{attribute 'no_assign'}
FUNCTION_BLOCK FB_DO_WTURBINE_LD0_LPHD1_Proxy EXTENDS FB_AcsiCommonDataClass
VAR_INPUT
	stVal: FB_AcsiBATypeBOOLEAN := (Fc:=ACSI_FC_ST, TrgOp:=ACSI_TrgOp_dchg, bLinkResult:=THIS^.AddDataToContainer(ipData:=stVal));
	q: FB_AcsiDATypeQuality := (Fc:=ACSI_FC_ST, TrgOp:=ACSI_TrgOp_qchg, bLinkResult:=THIS^.AddDataToContainer(ipData:=q));
	t: FB_AcsiDATypeTimeStamp := (Fc:=ACSI_FC_ST, bLinkResult:=THIS^.AddDataToContainer(ipData:=t));
END_VAR
VAR
END_VAR

END_FUNCTION_BLOCK

(* stored: Version 1.1.0.1
   POU FB_DO_WTURBINE_LD0_LPHD1_Proxy: Id {51a2d004-d7e3-4470-9c80-0b470bf52205}, SpecialFunc None *)
